(* IEC 61131-3 sources: rusty/tests/lit/multi/direct_linker_shared, 1 file *)

(* ---- add_one.st ---- *)
FUNCTION addOne : DINT
VAR_INPUT
    value : DINT;
END_VAR
    addOne := value + 1;
END_FUNCTION
